(* IEC 61131-3 sources: Lasal-MCP/examples/SampleSource/4_PumpControlSchemeSolution/Stations/MachineControl/MachineControl/Class/PumpControlSimu, 1 file *)

(* ---- PumpControlSimu.st ---- *)
(*!
<Class
	Name               = "PumpControlSimu"
	Revision           = "0.0"
	RealtimeTask       = "false"
	DefRealtime        = "1 ms"
	CyclicTask         = "true"
	DefCyclictime      = "1 ms"
	BackgroundTask     = "false"
	Sigmatek           = "false"
	OSInterface        = "false"
	HighPriority       = "false"
	Automatic          = "false"
	UpdateMode         = "Prescan"
	SharedCommandTable = "true"
	Objectsize         = "(380,120)">
	<Channels>
		<Server Name="FillLevel" Visualized="false" Initialize="false" WriteProtected="true" Retentive="false"/>
		<Server Name="Pump" Visualized="false" Initialize="false" WriteProtected="false" Retentive="false"/>
		<Server Name="SimuSpeed" Visualized="true" Initialize="false" WriteProtected="false" Retentive="File"/>
		<Server Name="SimuStart" Visualized="true" Initialize="false" WriteProtected="false" Retentive="false"/>
		<Server Name="WaterTemp" Visualized="false" Initialize="false" WriteProtected="true" Retentive="false"/>
	</Channels>
</Class>
*)
PumpControlSimu : CLASS
  //Servers:
	FillLevel 	: SvrChCmd_DINT;
	Pump 	: SvrCh_DINT;
	WaterTemp 	: SvrCh_DINT;
	SimuSpeed 	: SvrCh_DINT;
	SimuStart 	: SvrCh_DINT;
  //Clients:
  //Variables:
		countup 	: DINT;
  //Functions:

	FUNCTION VIRTUAL GLOBAL Init;

	FUNCTION VIRTUAL GLOBAL CyWork
		VAR_INPUT
			EAX 	: UDINT;
		END_VAR
		VAR_OUTPUT
			state (EAX) 	: UDINT;
		END_VAR;
  //Tables:
	FUNCTION @STD
		VAR_OUTPUT
			ret_code	: CONFSTATES;
		END_VAR;
	FUNCTION GLOBAL TAB @CT_;
END_CLASS;

FUNCTION VIRTUAL GLOBAL PumpControlSimu::Init

  if _FirstScan then
    WaterTemp := 245;
  end_if;

END_FUNCTION

FUNCTION VIRTUAL GLOBAL PumpControlSimu::CyWork
	VAR_INPUT
		EAX 	: UDINT;
	END_VAR
	VAR_OUTPUT
		state (EAX) 	: UDINT;
	END_VAR

  if SimuStart = 1 then  // Start/Stop Simu

    if FillLevel = 0 | Pump = 0 then
       countup := 1;  // Pump inactive -> Count up
    elsif FillLevel >= 50000 | Pump = 1 then
       countup := 0;  // Pump active -> Count down
    end_if;

    if countup = 1 | Pump = 0 then
      FillLevel += SimuSpeed; // Count up
    else
      FillLevel -= SimuSpeed; // Count down
    end_if;
  end_if;

	state := READY;

END_FUNCTION
